(* IEC 61131-3 sources: Lasal-MCP/examples/SampleSource/4_PumpControlSchemeSolution/Stations/Terminal/HMI/Class/_EventQueue, 1 file *)

(* ---- _EventQueue.st ---- *)
#define     EventQueue_MaxEntries     50

(*!
<Class
	Name               = "_EventQueue"
	Revision           = "1.7"
	RealtimeTask       = "false"
	CyclicTask         = "false"
	BackgroundTask     = "true"
	DefBackground      = "10 ms"
	Sigmatek           = "true"
	OSInterface        = "false"
	HighPriority       = "false"
	Automatic          = "false"
	UpdateMode         = "Prescan"
	SharedCommandTable = "true"
	Objectsize         = "(540,480)"
	Comment            = "class for converting row events and buffering for the EventJournal ">
	<Channels>
		<Server Name="ActEntries" Visualized="false" Initialize="false" WriteProtected="true" Retentive="false" Comment="actual number of entries in buffer to be readed/handled"/>
		<Server
			Name           = "ClassSvr"
			Visualized     = "false"
			Initialize     = "false"
			WriteProtected = "true"
			Retentive      = "false"
			Comment        = "class server">
			<NewInst>
				<Function Name="NewInst_AddSystemOnOff" Comment="AddSystemOnOff() via command channel">
					<InputParameter>
						<Parameter Name="dDate"/>
						<Parameter Name="dTime"/>
						<Parameter Name="bSwitchOnOff"/>
					</InputParameter>
					<OutputParameter>
						<Parameter Name="ret_code"/>
					</OutputParameter>
				</Function>
				<Function Name="NewInst_AddEventEntry" Comment="AddEventEntry() via command channel">
					<InputParameter>
						<Parameter Name="config"/>
						<Parameter Name="uiCategory"/>
						<Parameter Name="uiIndex"/>
						<Parameter Name="dParam1"/>
						<Parameter Name="pText"/>
						<Parameter Name="bUnicode"/>
					</InputParameter>
					<OutputParameter>
						<Parameter Name="ret_code"/>
					</OutputParameter>
				</Function>
				<Function Name="NewInst_AddDateChange" Comment="AddDateChange() via command channel">
					<InputParameter>
						<Parameter Name="udVarNo"/>
						<Parameter Name="dOldDate"/>
						<Parameter Name="dNewDate"/>
					</InputParameter>
					<OutputParameter>
						<Parameter Name="ret_code"/>
					</OutputParameter>
				</Function>
				<Function Name="NewInst_AddTimeChange" Comment="AddTimeChange() via command channel">
					<InputParameter>
						<Parameter Name="udVarNo"/>
						<Parameter Name="dOldTime"/>
						<Parameter Name="dNewTime"/>
					</InputParameter>
					<OutputParameter>
						<Parameter Name="ret_code"/>
					</OutputParameter>
				</Function>
				<Function Name="NewInst_AddMenuChange" Comment="AddMenuChange() via command channel">
					<InputParameter>
						<Parameter Name="udVarNo"/>
						<Parameter Name="udMenuIndex"/>
						<Parameter Name="dOldValue"/>
						<Parameter Name="dNewValue"/>
					</InputParameter>
					<OutputParameter>
						<Parameter Name="ret_code"/>
					</OutputParameter>
				</Function>
				<Function Name="NewInst_AddValueChange" Comment="AddValueChange() via command channel">
					<InputParameter>
						<Parameter Name="udVarNo"/>
						<Parameter Name="dOldValue"/>
						<Parameter Name="dNewValue"/>
					</InputParameter>
					<OutputParameter>
						<Parameter Name="ret_code"/>
					</OutputParameter>
				</Function>
				<Function Name="NewInst_AddOPChange" Comment="AddOPChange() via command channel">
					<InputParameter>
						<Parameter Name="eOPMode"/>
					</InputParameter>
					<OutputParameter>
						<Parameter Name="ret_code"/>
					</OutputParameter>
				</Function>
				<Function Name="NewInst_AddUserLoginLogout">
					<InputParameter>
						<Parameter Name="pUserName"/>
						<Parameter Name="dActLevel"/>
						<Parameter Name="bIsLogin"/>
					</InputParameter>
					<OutputParameter>
						<Parameter Name="ret_code"/>
					</OutputParameter>
				</Function>
			</NewInst>
		</Server>
		<Server Name="MaxEntries" Visualized="false" Initialize="false" WriteProtected="true" Retentive="false" Comment="max. number of entries in buffer to be readed/handled"/>
		<Client Name="ccSystemLogging" Required="false" Internal="false" Comment="command channel to SystemLogging (optional)"/>
		<Client Name="coEventJournal" Required="true" Internal="false" Comment="object channel to EventJournal"/>
		<Client Name="coGraphic" Required="false" Internal="false" Comment="object channel to Graphic (don&apos;t connect!)"/>
		<Client Name="coStdLib" Required="false" Internal="false" Comment="object channel to SdtLib (don&apos;t connect!)"/>
		<Client Name="Param1" Required="true" Internal="false" Comment="Parameter 1 for event entry"/>
		<Client Name="Param2" Required="true" Internal="false" Comment="Parameter 2 for event entry"/>
		<Client Name="SysDate" Required="true" Internal="false" Comment="object channel to SysDate"/>
		<Client Name="SysTime" Required="true" Internal="false" Comment="object channel to SysTime"/>
	</Channels>
	<Dependencies>
		<Files>
			<File Path=".\Class\_EventJournal\Event.h" Include="true"/>
			<File Path=".\Class\_EventQueue\_EventQueue_de.pdf"/>
			<File Path=".\Class\_EventQueue\_EventQueue_en.pdf"/>
		</Files>
	</Dependencies>
	<RevDoku>
		<Owner Company="Sigmatek"/>
		<Dokumentation Revision="1.7" Date="2016-10-10" Author="HubChr" Company="Sigmatek" Description="Added documentation pdfs."/>
		<Dokumentation Revision="1.6" Date="2016-10-06" Author="KaiAnd" Company="Sigmatek" Description="implemented NewInst_AddXY (Cmd 00 to Cmd 07) for adding events from external via command channel"/>
		<Dokumentation Revision="1.5" Date="2016-09-29" Author="KaiAnd" Company="Sigmatek" Description="changed object channel for SystemLogging to a command channel; new help function LogMyText() for logging"/>
		<Dokumentation Revision="1.4" Date="2016-09-19" Author="KaiAnd" Company="Sigmatek" Description="--&gt; ::AddEventEntry() got a new input &quot;dParam1&quot; as parameter 1 for the event &#13;&#10;... if this value is #0 the value of the client &quot;Param1&quot; will be used&#13;&#10;--&gt; ::AddEventEntry() got a new input &quot;config&quot; with event configuration bits&#13;&#10;... Bit 0:  1= add event to EventJournal / Bit 1:  1= create a MessageBox&#13;&#10;... the creation of the message box will happen here"/>
		<Dokumentation Revision="1.3" Date="2016-08-22" Author="Roskri" Company="Sigmatek" Description="Clients SysDate and SysTime changed to HDINT"/>
		<Dokumentation Revision="1.2" Date="2016-05-18" Author="KaiAnd" Company="Sigmatek" Description="object channel to SystemLogging is optional now"/>
		<Dokumentation Revision="1.1" Date="2015-05-22" Author="BraLis" Company="Sigmatek" Description="insert the method SystemLogging::LogEventText instead of TRACE-Messages"/>
		<Dokumentation Revision="1.0" Date="2015-03-31" Company="Sigmatek" Description="Creation&#13;&#10;"/>
	</RevDoku>
</Class>
*)
_EventQueue : CLASS
	TYPE
	  CmdClassSvr :  //! <Type Public="true" Name="CmdClassSvr"/>
	  (
	    NewInst_AddSystemOnOff,
	    NewInst_AddEventEntry,
	    NewInst_AddDateChange,
	    NewInst_AddTimeChange,
	    NewInst_AddMenuChange,
	    NewInst_AddValueChange,
	    NewInst_AddOPChange,
	    NewInst_AddUserLoginLogout
	  )$UINT;
#pragma pack(push, 1)
	  t_s_EventBuffer : STRUCT
	    pStart : ^_SINGLEALARM;
	    pEnd : ^_SINGLEALARM;
	    pWrite : ^_SINGLEALARM;
	    pRead : ^_SINGLEALARM;
	    udSize : UDINT;
	    udElements : UDINT;
	  END_STRUCT;
#pragma pack(pop)
	END_TYPE
  //Servers:
	ClassSvr 	: SvrChCmd_DINT;
	ActEntries 	: SvrCh_UDINT;
	MaxEntries 	: SvrCh_UDINT;
  //Clients:
	coGraphic 	: CltChCmd_Graphic;
	coEventJournal 	: CltChCmd__EventJournal;
	Param1 	: CltCh_DINT;
	Param2 	: CltCh_DINT;
	SysDate 	: CltCh_HDINT;
	SysTime 	: CltCh_HDINT;
	coStdLib 	: CltChCmd__StdLib;
	ccSystemLogging 	: CltChCmd_DINT;
  //Variables:
		sEventBuffer 	: t_s_EventBuffer;
		IsCon_ccSystemLogging 	: BOOL;
		MsgBoxInit 	: DINT;			//! <Variable Comment="INIT for message boxes is necessary" Name="MsgBoxInit"/>
  //Functions:

	FUNCTION VIRTUAL GLOBAL Init;

	FUNCTION VIRTUAL GLOBAL Background
		VAR_INPUT
			EAX 	: UDINT;
		END_VAR
		VAR_OUTPUT
			state (EAX) 	: UDINT;
		END_VAR;
				//! <Function Comment="This Method is used to register an event into the logbook." Name="AddEventEntry"/>
	FUNCTION GLOBAL AddEventEntry
		VAR_INPUT
			config 	: BDINT;			//! <Variable Comment="configuration bits&#13;&#10;Bit 0:  1= add event to EventJournal&#13;&#10;Bit 1:  1= create a MessageBox" Name="AddEventEntry.config"/>
			uiCategory 	: UINT;			//! <Variable Comment="Category for the event:&#13;&#10;0 .. System category 1&#13;&#10;1 .. System category 2&#13;&#10;2 .. System category 3&#13;&#10;3 .. System category 4&#13;&#10;4 .. Change of the OP mode&#13;&#10;else .. System category 1" Name="AddEventEntry.uiCategory"/>
			uiIndex 	: UINT;			//! <Variable Comment="Index in the textscheme (if used).&#13;&#10;Note: If event is for example a menue-change -&gt; menue-index." Name="AddEventEntry.uiIndex"/>
			dParam1 	: DINT;			//! <Variable Comment="parameter 1 for the event &#13;&#10;... if this value is #0 the value of the client &quot;Param1&quot; will be used" Name="AddEventEntry.dParam1"/>
			pText 	: ^void;			//! <Variable Comment="Individual text" Name="AddEventEntry.pText"/>
			bUnicode 	: BOOL;			//! <Variable Comment="Character size of the string:&#13;&#10;FALSE .. ASCII&#13;&#10;TRUE .. UNI-Code" Name="AddEventEntry.bUnicode"/>
		END_VAR
		VAR_OUTPUT
			bSuccessful 	: BOOL;			//! <Variable Comment="FALSE..Event could not be inserted into the buffer&#13;&#10;TRUE..Event inserted successfullly" Name="AddEventEntry.bSuccessful"/>
		END_VAR;
				//! <Function Comment="Method to insert an event for a date change into the buffer." Name="AddDateChange"/>
	FUNCTION GLOBAL AddDateChange
		VAR_INPUT
			udVarNo 	: UDINT;			//! <Variable Comment="Variable number" Name="AddDateChange.udVarNo"/>
			dOldDate 	: DINT;			//! <Variable Comment="Old date" Name="AddDateChange.dOldDate"/>
			dNewDate 	: DINT;			//! <Variable Comment="New date" Name="AddDateChange.dNewDate"/>
		END_VAR
		VAR_OUTPUT
			bSuccessful 	: BOOL;			//! <Variable Comment="FALSE..event could not be inserted into the buffer&#13;&#10;TRUE..event inserted successfully" Name="AddDateChange.bSuccessful"/>
		END_VAR;
				//! <Function Comment="Method to insert an event for a time change into the buffer" Name="AddTimeChange"/>
	FUNCTION GLOBAL AddTimeChange
		VAR_INPUT
			udVarNo 	: UDINT;			//! <Variable Comment="Variable number" Name="AddTimeChange.udVarNo"/>
			dOldTime 	: DINT;			//! <Variable Comment="Old time" Name="AddTimeChange.dOldTime"/>
			dNewTime 	: DINT;			//! <Variable Comment="New time" Name="AddTimeChange.dNewTime"/>
		END_VAR
		VAR_OUTPUT
			bSuccessful 	: BOOL;			//! <Variable Comment="FALSE..Event could not be inserted to the buffer&#13;&#10;TRUE..Event inserted successfully" Name="AddTimeChange.bSuccessful"/>
		END_VAR;
				//! <Function Comment="Method to insert an event for a menu change into the buffer." Name="AddMenuChange"/>
	FUNCTION GLOBAL AddMenuChange
		VAR_INPUT
			udVarNo 	: UDINT;			//! <Variable Comment="Variable number" Name="AddMenuChange.udVarNo"/>
			udMenuIndex 	: UDINT;
			dOldValue 	: DINT;			//! <Variable Comment="Old value" Name="AddMenuChange.dOldValue"/>
			dNewValue 	: DINT;			//! <Variable Comment="New value" Name="AddMenuChange.dNewValue"/>
		END_VAR
		VAR_OUTPUT
			bSuccessful 	: BOOL;			//! <Variable Comment="FALSE..Event could not be inserted into the buffer&#13;&#10;TRUE..Event inserted successfully" Name="AddMenuChange.bSuccessful"/>
		END_VAR;
				//! <Function Comment="Method to insert an event for a value change into the buffer." Name="AddValueChange"/>
	FUNCTION GLOBAL AddValueChange
		VAR_INPUT
			udVarNo 	: UDINT;			//! <Variable Comment="Variable number" Name="AddValueChange.udVarNo"/>
			dOldValue 	: DINT;			//! <Variable Comment="Old value" Name="AddValueChange.dOldValue"/>
			dNewValue 	: DINT;			//! <Variable Comment="New value" Name="AddValueChange.dNewValue"/>
		END_VAR
		VAR_OUTPUT
			bSuccessful 	: BOOL;			//! <Variable Comment="FALSE..Event could not be inserted into the buffer&#13;&#10;TRUE..Event inserted successfully" Name="AddValueChange.bSuccessful"/>
		END_VAR;
				//! <Function Comment="Method to insert an event for the change of the operation mode into the buffer." Name="AddOPChange"/>
	FUNCTION GLOBAL AddOPChange
		VAR_INPUT
			eOPMode 	: t_e_OPMode;			//! <Variable Comment="New operation mode" Name="AddOPChange.eOPMode"/>
		END_VAR
		VAR_OUTPUT
			bSuccessful 	: BOOL;			//! <Variable Comment="FALSE..Event could not be insert into the buffer&#13;&#10;TRUE..Event inserted successfully" Name="AddOPChange.bSuccessful"/>
		END_VAR;
				//! <Function Comment="Method to insert an event for turning on or off the system." Name="AddSystemOnOff"/>
	FUNCTION VIRTUAL GLOBAL AddSystemOnOff
		VAR_INPUT
			dDate 	: DINT;			//! <Variable Comment="Actual date" Name="AddSystemOnOff.dDate"/>
			dTime 	: DINT;			//! <Variable Comment="Actual time" Name="AddSystemOnOff.dTime"/>
			bSwitchOnOff 	: BOOL;			//! <Variable Comment="FALSE..Event for turning off the system&#13;&#10;TRUE..Event for turning on the system" Name="AddSystemOnOff.bSwitchOnOff"/>
		END_VAR
		VAR_OUTPUT
			bSuccessful 	: BOOL;			//! <Variable Comment="FALSE..Event could not be inserted to the buffer&#13;&#10;TRUE..Event inserted succesfully" Name="AddSystemOnOff.bSuccessful"/>
		END_VAR;
				//! <Function Comment="Method to insert an user event (text) into the buffer" Name="AddUserEvent"/>
	FUNCTION GLOBAL AddUserEvent
		VAR_INPUT
			pEventString 	: ^_CHAR;			//! <Variable Comment="Pointer to the text which should be added (Unicode)" Name="AddUserEvent.pEventString"/>
		END_VAR
		VAR_OUTPUT
			bSuccessful 	: BOOL;			//! <Variable Comment="FALSE..Event could not be inserted into the buffer&#13;&#10;TRUE..Event inserted successfully" Name="AddUserEvent.bSuccessful"/>
		END_VAR;
				//! <Function Comment="Method to insert an event for user login/logout into the buffer." Name="AddUserLoginLogout"/>
	FUNCTION GLOBAL AddUserLoginLogout
		VAR_INPUT
			pUserName 	: ^CHAR;			//! <Variable Comment="Pointer to the name of the user, which was logged in or logged out" Name="AddUserLoginLogout.pUserName"/>
			dActLevel 	: DINT;			//! <Variable Comment="User level" Name="AddUserLoginLogout.dActLevel"/>
			bIsLogin 	: BOOL;			//! <Variable Comment="FALSE..User logged out&#13;&#10;TRUE..User logged in" Name="AddUserLoginLogout.bIsLogin"/>
		END_VAR
		VAR_OUTPUT
			bSuccessful 	: BOOL;			//! <Variable Comment="FALSE..Event could not be inserted to the buffer&#13;&#10;TRUE..Event inserted successfully" Name="AddUserLoginLogout.bSuccessful"/>
		END_VAR;
				//! <Function Comment="Copy data into the write buffer and set the write pointer so that the entry in the buffer will be added to the event journal in the next background run." Name="AddEntry"/>
	FUNCTION AddEntry
		VAR_INPUT
			pEntry 	: ^_SINGLEALARM;			//! <Variable Comment="Pointer to the data of the entry" Name="AddEntry.pEntry"/>
		END_VAR
		VAR_OUTPUT
			bSuccessful 	: BOOL;			//! <Variable Comment="FALSE..pEntry was NIL&#13;&#10;TRUE..Ok" Name="AddEntry.bSuccessful"/>
		END_VAR;
				//! <Function Comment="help function to log a text via command channel to SystemLogging" Name="LogMyText"/>
	FUNCTION LogMyText
		VAR_INPUT
			pLogTxt 	: ^CHAR;			//! <Variable Comment="pointer to the text which should be logged" Name="LogMyText.pLogTxt"/>
		END_VAR;
				//! <Function Comment="AddSystemOnOff() via command channel" Name="ClassSvr.NewInst_AddSystemOnOff"/>
	FUNCTION ClassSvr::NewInst_AddSystemOnOff
		VAR_INPUT
			dDate 	: DINT;
			dTime 	: DINT;
			bSwitchOnOff 	: DINT;
		END_VAR
		VAR_OUTPUT
			ret_code 	: IprStates;
		END_VAR;
				//! <Function Comment="AddEventEntry() via command channel" Name="ClassSvr.NewInst_AddEventEntry"/>
	FUNCTION ClassSvr::NewInst_AddEventEntry
		VAR_INPUT
			config 	: DINT;
			uiCategory 	: DINT;
			uiIndex 	: DINT;
			dParam1 	: DINT;
			pText 	: DINT;
			bUnicode 	: DINT;
		END_VAR
		VAR_OUTPUT
			ret_code 	: IprStates;
		END_VAR;
				//! <Function Comment="AddDateChange() via command channel" Name="ClassSvr.NewInst_AddDateChange"/>
	FUNCTION ClassSvr::NewInst_AddDateChange
		VAR_INPUT
			udVarNo 	: DINT;
			dOldDate 	: DINT;
			dNewDate 	: DINT;
		END_VAR
		VAR_OUTPUT
			ret_code 	: IprStates;
		END_VAR;
				//! <Function Comment="AddTimeChange() via command channel" Name="ClassSvr.NewInst_AddTimeChange"/>
	FUNCTION ClassSvr::NewInst_AddTimeChange
		VAR_INPUT
			udVarNo 	: DINT;
			dOldTime 	: DINT;
			dNewTime 	: DINT;
		END_VAR
		VAR_OUTPUT
			ret_code 	: IprStates;
		END_VAR;
				//! <Function Comment="AddMenuChange() via command channel" Name="ClassSvr.NewInst_AddMenuChange"/>
	FUNCTION ClassSvr::NewInst_AddMenuChange
		VAR_INPUT
			udVarNo 	: DINT;
			udMenuIndex 	: DINT;
			dOldValue 	: DINT;
			dNewValue 	: DINT;
		END_VAR
		VAR_OUTPUT
			ret_code 	: IprStates;
		END_VAR;
				//! <Function Comment="AddValueChange() via command channel" Name="ClassSvr.NewInst_AddValueChange"/>
	FUNCTION ClassSvr::NewInst_AddValueChange
		VAR_INPUT
			udVarNo 	: DINT;
			dOldValue 	: DINT;
			dNewValue 	: DINT;
		END_VAR
		VAR_OUTPUT
			ret_code 	: IprStates;
		END_VAR;
				//! <Function Comment="AddOPChange() via command channel" Name="ClassSvr.NewInst_AddOPChange"/>
	FUNCTION ClassSvr::NewInst_AddOPChange
		VAR_INPUT
			eOPMode 	: DINT;
		END_VAR
		VAR_OUTPUT
			ret_code 	: IprStates;
		END_VAR;

	FUNCTION ClassSvr::NewInst_AddUserLoginLogout
		VAR_INPUT
			pUserName 	: DINT;
			dActLevel 	: DINT;
			bIsLogin 	: DINT;
		END_VAR
		VAR_OUTPUT
			ret_code 	: IprStates;
		END_VAR;
				//! <Function Name="ClassSvr.NewInst" Hidden="true"/>
	FUNCTION VIRTUAL GLOBAL ClassSvr::NewInst
		VAR_INPUT
			pPara 	: ^CmdStruct;
			pResult 	: ^results;
		END_VAR
		VAR_OUTPUT
			ret_code 	: iprStates;
		END_VAR;
  //Tables:
	FUNCTION @STD
		VAR_OUTPUT
			ret_code	: CONFSTATES;
		END_VAR;
	FUNCTION GLOBAL TAB @CT_;
END_CLASS;

#pragma usingLtd _EventJournal
#pragma usingLtd _StdLib
#pragma usingLtd Graphic

FUNCTION VIRTUAL GLOBAL _EventQueue::ClassSvr::NewInst
	VAR_INPUT
		pPara 	: ^CmdStruct;
		pResult 	: ^Results;
	END_VAR
	VAR_OUTPUT
		ret_code 	: IprStates;
	END_VAR
	CASE pPara^.uiCmd$CmdClassSvr OF
		NewInst_AddSystemOnOff:
			ret_code := NewInst_AddSystemOnOff(pPara^.aPara[0],pPara^.aPara[1],pPara^.aPara[2]);
			pResult^.uiLng := 0 + sizeof(pResult^.uiLng);
		NewInst_AddEventEntry:
			ret_code := NewInst_AddEventEntry(pPara^.aPara[0],pPara^.aPara[1],pPara^.aPara[2],pPara^.aPara[3],pPara^.aPara[4],pPara^.aPara[5]);
			pResult^.uiLng := 0 + sizeof(pResult^.uiLng);
		NewInst_AddDateChange:
			ret_code := NewInst_AddDateChange(pPara^.aPara[0],pPara^.aPara[1],pPara^.aPara[2]);
			pResult^.uiLng := 0 + sizeof(pResult^.uiLng);
		NewInst_AddTimeChange:
			ret_code := NewInst_AddTimeChange(pPara^.aPara[0],pPara^.aPara[1],pPara^.aPara[2]);
			pResult^.uiLng := 0 + sizeof(pResult^.uiLng);
		NewInst_AddMenuChange:
			ret_code := NewInst_AddMenuChange(pPara^.aPara[0],pPara^.aPara[1],pPara^.aPara[2],pPara^.aPara[3]);
			pResult^.uiLng := 0 + sizeof(pResult^.uiLng);
		NewInst_AddValueChange:
			ret_code := NewInst_AddValueChange(pPara^.aPara[0],pPara^.aPara[1],pPara^.aPara[2]);
			pResult^.uiLng := 0 + sizeof(pResult^.uiLng);
		NewInst_AddOPChange:
			ret_code := NewInst_AddOPChange(pPara^.aPara[0]);
			pResult^.uiLng := 0 + sizeof(pResult^.uiLng);
		NewInst_AddUserLoginLogout:
			ret_code := NewInst_AddUserLoginLogout(pPara^.aPara[0],pPara^.aPara[1],pPara^.aPara[2]);
			pResult^.uiLng := 0 + sizeof(pResult^.uiLng);
	ELSE

	ret_code := READY;
	END_CASE;

END_FUNCTION

FUNCTION VIRTUAL GLOBAL _EventQueue::Init
VAR
	tmpMemory : ^_SINGLEALARM;
END_VAR

  // letzter Init-Durchlauf
  if (_FirstScan) then

    //-------------------------------------------------------------------------
    //  check client-connnections and set flags		KaiAnd
    //-------------------------------------------------------------------------
    if (IsClientConnected(#ccSystemLogging)) then
      IsCon_ccSystemLogging := TRUE;
    else
      IsCon_ccSystemLogging := FALSE;
    end_if;

    MsgBoxInit := TRUE;   // INIT for message boxes is necessary  V.1.4, KaiAnd

    // Speicher für Eventbuffer allokieren
    tmpMemory$^void := coStdLib.Malloc(size := EventQueue_MaxEntries * sizeof(sEventBuffer.pStart^));

    // Prüfen ob Speicher verfügbar
    if (tmpMemory <> NIL) then

      // Größe vom Buffer speichern
      sEventBuffer.udElements := EventQueue_MaxEntries;
      sEventBuffer.udSize     := EventQueue_MaxEntries * sizeof(sEventBuffer.pStart^);

      // Pointer für Buffer speichern
      sEventBuffer.pStart := tmpMemory;
      sEventBuffer.pEnd   := tmpMemory + sEventBuffer.udSize;
      sEventBuffer.pRead  := tmpMemory;
      sEventBuffer.pWrite := tmpMemory;

    else
      LogMyText("_EventQueue::Init(): allokieren des Eventspeichers fehlgeschlagen");
    end_if;

  end_if;

END_FUNCTION

FUNCTION VIRTUAL GLOBAL _EventQueue::Background
	VAR_INPUT
		EAX 	: UDINT;
	END_VAR
	VAR_OUTPUT
		state (EAX) 	: UDINT;
	END_VAR

  // aktuelle Anzahl der Elemente im Buffer darstellen
  if (sEventBuffer.pWrite >= sEventBuffer.pRead) then
    ActEntries := (sEventBuffer.pWrite$UDINT - sEventBuffer.pRead$UDINT) / sizeof(sEventBuffer.pWrite^);
  else
    ActEntries := ((sEventBuffer.pEnd$UDINT - sEventBuffer.pRead$UDINT) + (sEventBuffer.pWrite$UDINT - sEventBuffer.pStart$UDINT)) / sizeof(sEventBuffer.pWrite^);
  end_if;

  // maximale Anzahl der Einträge darstellen
  if (ActEntries > MaxEntries) then
    MaxEntries := ActEntries;

    if (MaxEntries >= sEventBuffer.udElements -1) then
      LogMyText("_EventQueue::Background(): Bufferüberlauf");
    end_if;

  end_if;

  //*****************************************************************************
  //** SCHLEIFE ZUM LEEREN VOM BUFFER                                          **
  //*****************************************************************************
  while (sEventBuffer.pRead <> sEventBuffer.pWrite) do

    // Event an _EventJournal weiterleiten
    if (coEventJournal.AddEntry(ptr := sEventBuffer.pRead) = false) then
      LogMyText("_EventQueue::Background(): Eintragen des Events in _EventJournal fehlgeschlagen");
    end_if;

    // Auf nächsten Eintrag wechseln
    sEventBuffer.pRead += sizeof(sEventBuffer.pRead^);

    // Ende vom Buffer überwachen
    if (sEventBuffer.pRead >= sEventBuffer.pEnd) then
      sEventBuffer.pRead := sEventBuffer.pStart;
    end_if;

  end_while;

	state := READY;

END_FUNCTION

FUNCTION _EventQueue::AddEntry
	VAR_INPUT
		pEntry 	: ^_SINGLEALARM;
	END_VAR
	VAR_OUTPUT
		bSuccessful 	: BOOL;
	END_VAR

  // Übergabeparameter prüfen
  if (pEntry = NIL) then
    LogMyText("_EventQueue::AddEntry(): Übergabeparameter pEntry = NIL");
    bSuccessful := false;
    return;
  end_if;

  // Element in Buffer speichern
  _memcpy(ptr1  := sEventBuffer.pWrite,
          ptr2  := pEntry,
          cntr  := sizeof(sEventBuffer.pWrite^));

  // Schreibpointer weiterschalten
  sEventBuffer.pWrite += sizeof(sEventBuffer.pWrite^);

  // Ende vom Buffer überwachen
  if (sEventBuffer.pWrite >= sEventBuffer.pEnd) then
    sEventBuffer.pWrite := sEventBuffer.pStart;
  end_if;

  // alles erfolgreich
  bSuccessful := true;

END_FUNCTION

FUNCTION VIRTUAL GLOBAL _EventQueue::AddSystemOnOff
	VAR_INPUT
		dDate 	: DINT;
		dTime 	: DINT;
		bSwitchOnOff 	: BOOL;
	END_VAR
	VAR_OUTPUT
		bSuccessful 	: BOOL;
	END_VAR
  VAR
  	tmpEvent : _SINGLEALARM;
  END_VAR

  // Event initialisieren
  init_SINGLEALARM(#tmpEvent);

  if (bSwitchOnOff = false) then
    // Event für das Ausschalten der Steuerung
    tmpEvent.entrytype := EVENT_SWITCHOFF;
  else
    //Event für das Einschalten der Steuerung
    tmpEvent.entrytype := EVENT_SWITCHON;
  end_if;

  // Zyklusnummer lesen
  Param1 := Param1.Read();

  // Informationen speichern
  tmpEvent.no_para := 1;
  tmpEvent.para[0] := Param1;

  // Datum + Zeit speichern
  tmpEvent.date_on := dDate;
  tmpEvent.time_on := dTime;

  // Event zum Buffer hinzufügen
  if (AddEntry(pEntry := #tmpEvent) = true) then
    bSuccessful := true;
  else
    bSuccessful := false;
  end_if;

END_FUNCTION

FUNCTION GLOBAL _EventQueue::AddDateChange
	VAR_INPUT
		udVarNo 	: UDINT;
		dOldDate 	: DINT;
		dNewDate 	: DINT;
	END_VAR
	VAR_OUTPUT
		bSuccessful 	: BOOL;
	END_VAR
  VAR
  	tmpEvent : _SINGLEALARM;
  END_VAR

  // Event initialisieren
  init_SINGLEALARM(#tmpEvent);

  // Event für die Änderung eines Datums
  tmpEvent.entrytype := EVENT_DATECHANGE;

  // Zyklusnummer + Datum und Zeit + Zugangslevel lesen
  Param1  := Param1.Read();
  SysDate := SysDate.Read();
  SysTime := SysTime.Read();
  Param2  := Param2.Read();

  // Informationen speichern
  tmpEvent.no_para := 5;
  tmpEvent.para[0] := Param1;
  tmpEvent.para[1] := Param2;
  tmpEvent.para[2] := udVarNo$DINT;
  tmpEvent.para[3] := dOldDate;
  tmpEvent.para[4] := dNewDate;

  // Datum + Zeit speichern
  tmpEvent.date_on := to_dint(SysDate);
  tmpEvent.time_on := to_dint(SysTime);

  // Event zum Buffer hinzufügen
  if (AddEntry(pEntry := #tmpEvent) = true) then
    bSuccessful := true;
  else
    bSuccessful := false;
  end_if;

END_FUNCTION

FUNCTION GLOBAL _EventQueue::AddTimeChange
	VAR_INPUT
		udVarNo 	: UDINT;
		dOldTime 	: DINT;
		dNewTime 	: DINT;
	END_VAR
	VAR_OUTPUT
		bSuccessful 	: BOOL;
	END_VAR
  VAR
  	tmpEvent : _SINGLEALARM;
  END_VAR

  // Event initialisieren
  init_SINGLEALARM(#tmpEvent);

  // Event für die Änderung einer Zeit
  tmpEvent.entrytype := EVENT_TIMECHANGE;

  // Zyklusnummer + Datum und Zeit + Zugangslevel lesen
  Param1  := Param1.Read();
  SysDate := SysDate.Read();
  SysTime := SysTime.Read();
  Param2  := Param2.Read();

  // Informationen speichern
  tmpEvent.no_para := 5;
  tmpEvent.para[0] := Param1;
  tmpEvent.para[1] := Param2;
  tmpEvent.para[2] := udVarNo$DINT;
  tmpEvent.para[3] := dOldTime;
  tmpEvent.para[4] := dNewTime;

  // Datum + Zeit speichern
  tmpEvent.date_on := to_dint(SysDate);
  tmpEvent.time_on := to_dint(SysTime);

  // Event zum Buffer hinzufügen
  if (AddEntry(pEntry := #tmpEvent) = true) then
    bSuccessful := true;
  else
    bSuccessful := false;
  end_if;

END_FUNCTION

FUNCTION GLOBAL _EventQueue::AddValueChange
	VAR_INPUT
		udVarNo 	: UDINT;
		dOldValue 	: DINT;
		dNewValue 	: DINT;
	END_VAR
	VAR_OUTPUT
		bSuccessful 	: BOOL;
	END_VAR
  VAR
  	tmpEvent : _SINGLEALARM;
  END_VAR

  // Event initialisieren
  init_SINGLEALARM(#tmpEvent);

  // Event für die Änderung eines Wertes
  tmpEvent.entrytype := EVENT_VALUECHANGE;

  // Zyklusnummer + Datum und Zeit + Zugangslevel lesen
  Param1   := Param1.Read();
  SysDate  := SysDate.Read();
  SysTime  := SysTime.Read();
  Param2   := Param2.Read();

  // Informationen speichern
  tmpEvent.no_para := 5;
  tmpEvent.para[0] := Param1;
  tmpEvent.para[1] := Param2;
  tmpEvent.para[2] := udVarNo$DINT;
  tmpEvent.para[3] := dOldValue;
  tmpEvent.para[4] := dNewValue;

  // Datum + Zeit speichern
  tmpEvent.date_on := SysDate$DINT;
  tmpEvent.time_on := SysTime$DINT;

  // Event zum Buffer hinzufügen
  if (AddEntry(pEntry := #tmpEvent) = true) then
    bSuccessful := true;
  else
    bSuccessful := false;
  end_if;

END_FUNCTION

FUNCTION GLOBAL _EventQueue::AddMenuChange
	VAR_INPUT
		udVarNo 	: UDINT;
		udMenuIndex 	: UDINT;
		dOldValue 	: DINT;
		dNewValue 	: DINT;
	END_VAR
	VAR_OUTPUT
		bSuccessful 	: BOOL;
	END_VAR
  VAR
  	tmpEvent : _SINGLEALARM;
  END_VAR

  // Event initialisieren
  init_SINGLEALARM(#tmpEvent);

  // Event für die Änderung eines Wertes
  tmpEvent.entrytype := EVENT_MENUCHANGE;

  // Zyklusnummer + Datum und Zeit + Zugangslevel lesen
  Param1  := Param1.Read();
  SysDate := SysDate.Read();
  SysTime := SysTime.Read();
  Param2  := Param2.Read();

  // Informationen speichern
  tmpEvent.no_para := 6;
  tmpEvent.para[0] := Param1;
  tmpEvent.para[1] := Param2;
  tmpEvent.para[2] := udVarNo$DINT;
  tmpEvent.para[3] := dOldValue;
  tmpEvent.para[4] := dNewValue;
  tmpEvent.para[5] := udMenuIndex$DINT;

  // Datum + Zeit speichern
  tmpEvent.date_on := SysDate$DINT;
  tmpEvent.time_on := SysTime$DINT;

  // Event zum Buffer hinzufügen
  if (AddEntry(pEntry := #tmpEvent) = true) then
    bSuccessful := true;
  else
    bSuccessful := false;
  end_if;

END_FUNCTION

FUNCTION GLOBAL _EventQueue::AddOPChange
	VAR_INPUT
		eOPMode 	: t_e_OPMode;
	END_VAR
	VAR_OUTPUT
		bSuccessful 	: BOOL;
	END_VAR
  VAR
  	tmpEvent : _SINGLEALARM;
  END_VAR

  // Event initialisieren
  init_SINGLEALARM(#tmpEvent);

  // Event für die Änderung eines Wertes
  tmpEvent.entrytype := EVENT_OPCHANGE;

  // Zyklusnummer + Datum und Zeit + Zugangslevel lesen
  Param1  := Param1.Read();
  SysDate := SysDate.Read();
  SysTime := SysTime.Read();
  Param2  := Param2.Read();

  // Informationen speichern
  tmpEvent.no_para := 3;
  tmpEvent.para[0] := Param1;
  tmpEvent.para[1] := Param2;
  tmpEvent.para[2] := eOPMode$DINT;

  // Datum + Zeit speichern
  tmpEvent.date_on := SysDate$DINT;
  tmpEvent.time_on := SysTime$DINT;

  // Event zum Buffer hinzufügen
  if (AddEntry(pEntry := #tmpEvent) = true) then
    bSuccessful := true;
  else
    bSuccessful := false;
  end_if;

END_FUNCTION

FUNCTION GLOBAL _EventQueue::AddUserLoginLogout
	VAR_INPUT
		pUserName 	: ^CHAR;
		dActLevel 	: DINT;
		bIsLogin 	: BOOL;
	END_VAR
	VAR_OUTPUT
		bSuccessful 	: BOOL;
	END_VAR
  VAR
  	tmpEvent : _SINGLEALARM;
  END_VAR

  // Event initialisieren
  init_SINGLEALARM(#tmpEvent);

  if (bIsLogin = false) then
    tmpEvent.entrytype := Event_UserLogout;
  else
    tmpEvent.entrytype := Event_UserLogin;
  end_if;

  //Datum und Zeit lesen
  Param1  := Param1.Read();
  SysDate := SysDate.Read();
  SysTime := SysTime.Read();

  // Informationen speichern
  tmpEvent.no_para := 2;
  tmpEvent.para[0] := Param1;
  tmpEvent.para[1] := dActLevel;
  tmpEvent.ptrsize := (StrLen(txt:=pUserName, size:=sizeof(char)) + 1) * sizeof(_CHAR); // wegen Unicode
  tmpEvent.ptr     := coStdLib.Malloc(size:=tmpEvent.ptrsize);
  if (tmpEvent.ptr = NIL) then
    tmpEvent.ptrsize := 0;
    LogMyText("_EventQueue::AddUserLoginLogout(): Speicher für Benutzername konnte nicht reserviert werden");
  else
    StrCpy(p0:= tmpEvent.ptr, x1:= sizeof(_CHAR), p2:=pUserName, x3:=sizeof(CHAR));
  end_if;

  // Datum + Zeit speichern
  tmpEvent.date_on := SysDate$DINT;
  tmpEvent.time_on := SysTime$DINT;

  // Event zum Buffer hinzufügen
  if (AddEntry(pEntry := #tmpEvent) = true) then
    bSuccessful := true;
  else
    bSuccessful := false;
  end_if;

END_FUNCTION

FUNCTION GLOBAL _EventQueue::AddUserEvent
	VAR_INPUT
		pEventString 	: ^_CHAR;
	END_VAR
	VAR_OUTPUT
		bSuccessful 	: BOOL;
	END_VAR
  VAR
  	tmpEvent : _SINGLEALARM;
  END_VAR

  // Event initialisieren
  init_SINGLEALARM(#tmpEvent);

  // Event für die Änderung eines Wertes
  tmpEvent.entrytype := Event_UserEvent;

  // Zyklusnummer + Datum und Zeit + Zugangslevel lesen
  Param1  := Param1.Read();
  SysDate := SysDate.Read();
  SysTime := SysTime.Read();
  Param2  := Param2.Read();

  // Informationen speichern
  tmpEvent.no_para := 2;
  tmpEvent.para[0] := Param1;
  tmpEvent.para[1] := Param2;
  tmpEvent.ptrsize := sizeof(pEventString^) * (StrLen(txt:=pEventString, size:=sizeof(pEventString^)) + 1);
  tmpEvent.ptr     := coStdLib.Malloc(size:=tmpEvent.ptrsize);
  if (tmpEvent.ptr = NIL) then
    tmpEvent.ptrsize := 0;
    LogMyText("_EventQueue::AddUserEvent(): Speicher für Benutzer-Event konnte nicht reserviert werden");
  else
    _memcpy(ptr1:=tmpEvent.ptr, ptr2:=pEventString, cntr:=tmpEvent.ptrsize);
  end_if;

  // Datum + Zeit speichern
  tmpEvent.date_on := SysDate$DINT;
  tmpEvent.time_on := SysTime$DINT;

  // Event zum Buffer hinzufügen
  if (AddEntry(pEntry := #tmpEvent) = true) then
    bSuccessful := true;
  else
    bSuccessful := false;
  end_if;

END_FUNCTION

FUNCTION GLOBAL _EventQueue::AddEventEntry
	VAR_INPUT
		config 	: BDINT;
		uiCategory 	: UINT;
		uiIndex 	: UINT;
		dParam1 	: DINT;
		pText 	: ^void;
		bUnicode 	: BOOL;
	END_VAR
	VAR_OUTPUT
		bSuccessful 	: BOOL;
	END_VAR
  VAR
  	tmpEvent  :  _SINGLEALARM;
    pString   : ^_CHAR;
    actScreen : _NEWSCREEN;
    offScreen : _NEWSCREEN;
  END_VAR

  // Event initialisieren
  init_SINGLEALARM(#tmpEvent);
  bSuccessful := false;

  // Kategorie des Events definieren
  case (uiCategory) of
  0:
    tmpEvent.entrytype := Event_SystemCat1;
  1:
    tmpEvent.entrytype := Event_SystemCat2;
  2:
    tmpEvent.entrytype := Event_SystemCat3;
  3:
    tmpEvent.entrytype := Event_SystemCat4;
  4:
    tmpEvent.entrytype := Event_OPChange;
  else
    tmpEvent.entrytype := Event_SystemCat1;
  end_case;

  // Zyklusnummer + Datum und Zeit + Zugangslevel lesen
  Param1  := Param1.Read();
  SysDate := SysDate.Read();
  SysTime := SysTime.Read();
  Param2  := Param2.Read();

  // Informationen speichern
  tmpEvent.no_para := 3;
  if (dParam1 = 0) then         // V.1.4, KaiAnd use VAR_INPUT (dParam1) or client (Param1)
    tmpEvent.para[0] := Param1;
  else
    tmpEvent.para[0] := dParam1;
  end_if;
  tmpEvent.para[1] := Param2;
  tmpEvent.para[2] := uiIndex;

  // Speicher für den Text reservieren
  if (pText <> NIL) then

    if (bUnicode = true) then
      tmpEvent.ptrsize := (StrLen(txt:=pText, size:=sizeof(UINT)) + 1) * sizeof(UINT);
    else
      tmpEvent.ptrsize := (StrLen(txt:=pText, size:=sizeof(CHAR)) + 1) * sizeof(_CHAR);
    end_if;

    tmpEvent.ptr := coStdLib.Malloc(size:=tmpEvent.ptrsize);
    if (tmpEvent.ptr = NIL) then
      tmpEvent.ptrsize := 0;
      LogMyText("_EventQueue::AddEventEntry(): Speicher Eventtext konnte nicht reserviert werden");
    else

      if (bUnicode = true) then
        StrCpy(p0 := tmpEvent.ptr, x1 := sizeof(_CHAR), p2 := pText, x3 := sizeof(_CHAR));
      else
        StrCpy(p0 := tmpEvent.ptr, x1 := sizeof(_CHAR), p2 := pText, x3 := sizeof(CHAR));
      end_if;

    end_if;
  end_if;

  // Datum + Zeit speichern
  tmpEvent.date_on := SysDate$DINT;
  tmpEvent.time_on := SysTime$DINT;

  //-----------------------------------------------------------------------------------------------------
  //  ad Event to Buffer
  //  Config Bit 0: "add event to _EventJournal"  V.1.4, KaiAnd
  //-----------------------------------------------------------------------------------------------------
  if (config and 16#01) then
    if (AddEntry(pEntry := #tmpEvent) = true) then
      bSuccessful := true;
    else
      bSuccessful := false;
    end_if;
  end_if;

  //-----------------------------------------------------------------------------------------------------
  //  open a MessageBox ... V.1.4, KaiAnd
  //  Config Bit 1: "create a MessageBox"
  //-----------------------------------------------------------------------------------------------------
  if (config and 16#02) then

    //---------------------------------------------------------------------------------------------
    //  INIT for this message boxes
    //    this workarround is necessary because the _EventJournal must be opened 1 time to get
    //    the _EventJournal UDC-data - the _EventJournal need its UDC-data for GetEventText()
    //---------------------------------------------------------------------------------------------
    if (MsgBoxInit = TRUE) then
      if (coGraphic.CreateOffScreen(pScreen:=#offScreen, width:=100, height:=100)) then // create virtual OffScreen
        coGraphic.GetScreen(#actScreen);                // save the actual Screen
        coGraphic.SetScreen(#offScreen);                // switch to virtual OffScreen
        DrawPicWin(IMA_PICTURE, ScnNo_EventJournal, 5); // open the EbventJournal (into virtual offScreen)
        coGraphic.SetScreen( #actScreen);               // switch back to the saved actual screen
        coGraphic.DestroyOffScreen(#offScreen);         // kill the OffScreen
        free_NEWSCREEN(#offScreen);                     // free the offScreen memory
        MsgBoxInit := FALSE;                            // INIT done
      end_if;
    end_if;

    //---------------------------------------------------------------------------------------------
    //  open message box
    //---------------------------------------------------------------------------------------------
    pString := coEventJournal.GetEventText(#tmpEvent);

    MessageBoxSetFontScheme("Headline");

    MessageBoxSetFrame(box:=FRAME_WINDOW_NEWAGE, button:=FRAME_NEWAGE_DARK);

    MessageBoxSetColorBox(back  := coGraphic.MakeColor(MakeColorFromIndex(247), MakeColorFromIndex(242)),
                          text  := coGraphic.MakeColor(MakeColorFromIndex(246), MakeColorFromIndex(246)),
                          frame := coGraphic.MakeColor(MakeColorFromIndex(242), MakeColorFromIndex(242)) );

    MessageBoxSetColorButton(back  := coGraphic.MakeColor(MakeColorFromIndex(242), MakeColorFromIndex(242)),
                             text  := coGraphic.MakeColor(MakeColorFromIndex(241), MakeColorFromIndex(241)),
                             frame := coGraphic.MakeColor(MakeColorFromIndex(242), MakeColorFromIndex(242)) );

    MessageBoxCallEx(text:=pString, chrsize:=sizeof(_CHAR), typ:=MESSAGEBOXTYP_OK, pthis:=this, pfkt:=NIL);

    //---------------------------------------------------------------------------------------------

  end_if;
  //-----------------------------------------------------------------------------------------------------

END_FUNCTION

FUNCTION _EventQueue::LogMyText
  VAR_INPUT
		pLogTxt 	: ^CHAR;
	END_VAR

  VAR
    NiGive	  : CmdStruct;
    NiGet     : Results;
  END_VAR

  if ((IsCon_ccSystemLogging = True) & (pLogTxt <> NIL)) then

    NiGive.uiCmd    := 0;               // Command
    NiGive.aPara[0] := (pLogTxt)$DINT;  // pointer to text

    ccSystemLogging.NewInst(#NiGive, #NiGet);

  end_if;

END_FUNCTION

//***********************************************************************************************************
//  NewInst Commands for external actions via command channel
//***********************************************************************************************************

//-------------------------------------------------------------------------------------------------
//  Cmd 00: AddSystemOnOff
//-------------------------------------------------------------------------------------------------
FUNCTION _EventQueue::NewInst_AddSystemOnOff
	VAR_INPUT
		dDate 	: DINT;
		dTime 	: DINT;
		bSwitchOnOff 	: DINT;
	END_VAR
	VAR_OUTPUT
		ret_code 	: IprStates;
	END_VAR

	ret_code := READY;

  AddSystemOnOff( dDate        := dDate,
                  dTime        := dTime,
                  bSwitchOnOff := TO_BOOL(bSwitchOnOff) );

END_FUNCTION

//-------------------------------------------------------------------------------------------------
//  Cmd 01: AddEventEntry
//-------------------------------------------------------------------------------------------------
FUNCTION _EventQueue::NewInst_AddEventEntry
	VAR_INPUT
		config 	: DINT;
		uiCategory 	: DINT;
		uiIndex 	: DINT;
		dParam1 	: DINT;
		pText 	: DINT;
		bUnicode 	: DINT;
	END_VAR
	VAR_OUTPUT
		ret_code 	: IprStates;
	END_VAR

	ret_code := READY;

  AddEventEntry(config     := config$BDINT,
                uiCategory := TO_UINT(uiCategory),
                uiIndex    := TO_UINT(uiIndex),
                dParam1    := dParam1,
                pText      := pText$^void,
                bUnicode   := TO_BOOL(bUnicode) );

END_FUNCTION

//-------------------------------------------------------------------------------------------------
//  Cmd 02: AddDateChange
//-------------------------------------------------------------------------------------------------
FUNCTION _EventQueue::NewInst_AddDateChange
	VAR_INPUT
		udVarNo 	: DINT;
		dOldDate 	: DINT;
		dNewDate 	: DINT;
	END_VAR
	VAR_OUTPUT
		ret_code 	: IprStates;
	END_VAR

	ret_code := READY;

  AddDateChange(udVarNo  := udVarNo$UDINT,
                dOldDate := dOldDate,
                dNewDate := dNewDate );

END_FUNCTION

//-------------------------------------------------------------------------------------------------
//  Cmd 03: AddTimeChange
//-------------------------------------------------------------------------------------------------
FUNCTION _EventQueue::NewInst_AddTimeChange
	VAR_INPUT
		udVarNo 	: DINT;
		dOldTime 	: DINT;
		dNewTime 	: DINT;
	END_VAR
	VAR_OUTPUT
		ret_code 	: IprStates;
	END_VAR

	ret_code := READY;

  AddTimeChange(udVarNo  := udVarNo$UDINT,
                dOldTime := dOldTime,
                dNewTime := dNewTime );

END_FUNCTION

//-------------------------------------------------------------------------------------------------
//  Cmd 04: AddMenuChange
//-------------------------------------------------------------------------------------------------
FUNCTION _EventQueue::NewInst_AddMenuChange
	VAR_INPUT
		udVarNo 	: DINT;
		udMenuIndex 	: DINT;
		dOldValue 	: DINT;
		dNewValue 	: DINT;
	END_VAR
	VAR_OUTPUT
		ret_code 	: IprStates;
	END_VAR

	ret_code := READY;

  AddMenuChange(udVarNo     := udVarNo$UDINT,
                udMenuIndex := udMenuIndex$UDINT,
                dOldValue   := dOldValue,
                dNewValue   := dNewValue );

END_FUNCTION

//-------------------------------------------------------------------------------------------------
//  Cmd 05: AddValueChange
//-------------------------------------------------------------------------------------------------
FUNCTION _EventQueue::NewInst_AddValueChange
	VAR_INPUT
		udVarNo 	: DINT;
		dOldValue 	: DINT;
		dNewValue 	: DINT;
	END_VAR
	VAR_OUTPUT
		ret_code 	: IprStates;
	END_VAR

	ret_code := READY;

  AddValueChange( udVarNo   := udVarNo$UDINT,
                  dOldValue := dOldValue,
                  dNewValue := dNewValue );

END_FUNCTION

//-------------------------------------------------------------------------------------------------
//  Cmd 06: AddOPChange
//-------------------------------------------------------------------------------------------------
FUNCTION _EventQueue::NewInst_AddOPChange
	VAR_INPUT
		eOPMode 	: DINT;
	END_VAR
	VAR_OUTPUT
		ret_code 	: IprStates;
	END_VAR

	ret_code := READY;

  AddOPChange(eOPMode := eOPMode$t_e_OPMode);

END_FUNCTION

//-------------------------------------------------------------------------------------------------
//  Cmd 07: AddUserLoginLogout
//-------------------------------------------------------------------------------------------------
FUNCTION _EventQueue::NewInst_AddUserLoginLogout
	VAR_INPUT
		pUserName 	: DINT;
		dActLevel 	: DINT;
		bIsLogin 	: DINT;
	END_VAR
	VAR_OUTPUT
		ret_code 	: IprStates;
	END_VAR

	ret_code := READY;

  AddUserLoginLogout( pUserName := pUserName$^CHAR,
                      dActLevel := dActLevel,
                      bIsLogin  := TO_BOOL(bIsLogin) );

END_FUNCTION

//***********************************************************************************************************
